// Code-only delta: the interface and every DB remain unchanged.
FUNCTION "FC_S11RecoveryMarker" : Void
{ S7_Optimized_Access := 'TRUE' }
VERSION : 0.1
   VAR_IN_OUT
      Marker : DInt;
   END_VAR
BEGIN
    #Marker := 2101;
END_FUNCTION
